(* IEC 61131-3 sources: codesys-to-s7/tests/corpus/C2S7-SEM-CTR/neg, 1 file *)

(* ---- input.st ---- *)
FUNCTION_BLOCK FB_Case
VAR
    e : R_TRIG;
    x : BOOL;
END_VAR
e(CLK := x);
END_FUNCTION_BLOCK
